Fanuc KAREL source: KA00187.KL

PROGRAM KA00187
%NOLOCKGROUP
VAR
  SRC: ARRAY[4] OF BYTE
  DST: ARRAY[4] OF VECTOR
BEGIN
  DST = SRC
END KA00187
